Fanuc KAREL source: KD00047.KL

PROGRAM KD00047
%NOLOCKGROUP
%DEFGROUP = 1
VAR
  I: INTEGER
  J: INTEGER
  B: BOOLEAN
  R: REAL
  S: STRING[80]
  V: VECTOR
BEGIN
  V.X = 1.0
  MOVE ABOUT V BY 10.0
END KD00047
